// TwinCAT 3 PLC project BottleFactory
// ProgramVersion: 3.1.4026.28
// libraries:
//   CNM_AbstractObject, * (ekvip automation GmbH)
//   CNM_AssertionInterfaces, * (ekvip automation GmbH)
//   CNM_CommandInterfaces, * (ekvip automation GmbH)
//   CNM_CycleManager, * (ekvip automation GmbH)
//   CNM_CycleManagerInterfaces, * (ekvip automation GmbH)
//   CNM_MessageInterfaces, * (ekvip automation GmbH)
//   CNM_ReturnTypes, * (ekvip automation GmbH)
//   CNM_UnicodeUtilities, * (ekvip automation GmbH)
//   Tc2_Standard, * (Beckhoff Automation GmbH)
//   Tc2_System, * (Beckhoff Automation GmbH)
// project tree:
//   / PlcTask.TcTTO
//   POUs/ FB_CappingStation.TcPOU, FB_CinnamonFillingStation.TcPOU, FB_FillingStation.TcPOU, MAIN.TcPOU
// real-time tasks:
//   TASK PlcTask: cycle T#10ms, priority 20, ADS port 350

CONFIGURATION BottleFactory
    RESOURCE PLC ON TwinCAT3
        TASK PlcTask(INTERVAL := T#10ms, PRIORITY := 20);
        PROGRAM MAIN WITH PlcTask : MAIN;
    END_RESOURCE
END_CONFIGURATION

// ---- POUs/MAIN.TcPOU

PROGRAM MAIN
VAR
    bStart : BOOL := FALSE;
    bStop : BOOL := FALSE;
    bBottlePresent : BOOL := TRUE;

    fbStation : FB_FillingStation;
	fbCinnamon : FB_CinnamonFillingStation;
	bCinnamonRun : BOOL := FALSE;
	bCinnamonStop : BOOL := FALSE;
    nConveyorPosition : UDINT;
    nConveyorIndexBase : UDINT;
    nTransferPhase : UDINT;
    nPlaceProgress : UDINT;
    bBottleCapped : BOOL;
    fbInfeed : TON;
    fbOutfeed : TON;
    fbPlacement : TON;
    fbCapping : FB_CappingStation;
END_VAR


// 0: fill, 1: travel to capper, 2: cap, 3: pick and place, 4: bring next bottle to filler.
fbInfeed(IN := nTransferPhase = 1 AND NOT bCinnamonStop, PT := T#2S);
fbCapping(bBottleReady := nTransferPhase = 2, bStop := bCinnamonStop);
fbPlacement(IN := nTransferPhase = 3 AND NOT bCinnamonStop, PT := T#3S);
fbOutfeed(IN := nTransferPhase = 4 AND NOT bCinnamonStop, PT := T#2S);

IF NOT bCinnamonStop THEN
    CASE nTransferPhase OF
        0: IF fbCinnamon.bDone THEN nTransferPhase := 1; END_IF;
        1: IF fbInfeed.Q THEN nTransferPhase := 2; END_IF;
        2: IF fbCapping.bDone THEN nTransferPhase := 3; END_IF;
        3: IF fbPlacement.Q THEN nTransferPhase := 4; END_IF;
        4:
            IF fbOutfeed.Q THEN
                nConveyorIndexBase := nConveyorIndexBase + UDINT#100;
                nTransferPhase := 0;
            END_IF;
    END_CASE;

    nPlaceProgress := 0;
    nConveyorPosition := nConveyorIndexBase;
    CASE nTransferPhase OF
        1: nConveyorPosition := nConveyorIndexBase + DINT_TO_UDINT(TIME_TO_DINT(fbInfeed.ET) / DINT#40);
        2: nConveyorPosition := nConveyorIndexBase + UDINT#50;
        3:
            nConveyorPosition := nConveyorIndexBase + UDINT#50;
            nPlaceProgress := DINT_TO_UDINT(TIME_TO_DINT(fbPlacement.ET) / DINT#30);
        4:
            nConveyorPosition := nConveyorIndexBase + UDINT#50
                + DINT_TO_UDINT(TIME_TO_DINT(fbOutfeed.ET) / DINT#40);
            nPlaceProgress := 100;
    END_CASE;
END_IF;

bBottlePresent := nTransferPhase = 0;
bBottleCapped := nTransferPhase = 3;

fbStation(
    bStart := bStart,
    bStop := bStop,
    bBottlePresent := bBottlePresent
);


fbCinnamon(
    bRunRequest := bCinnamonRun,
    bStop := bCinnamonStop,
    bBottlePresent := bBottlePresent
);

END_PROGRAM

// ---- POUs/FB_FillingStation.TcPOU

FUNCTION_BLOCK FB_FillingStation
VAR_INPUT
    bStart : BOOL;
    bStop : BOOL;
    bBottlePresent : BOOL;
END_VAR

VAR_OUTPUT
    bValveOpen : BOOL;
    bBusy : BOOL;
    bDone : BOOL;
    nCompleted : UDINT;
END_VAR

VAR
    fbTimer : TON;
    fbStartEdge : R_TRIG;
    nState : INT := 0;
END_VAR


fbStartEdge(CLK := bStart);

fbTimer(
    IN := (nState = 10)
          AND NOT bStop
          AND bBottlePresent,
    PT := T#3S
);

bValveOpen := FALSE;
bBusy := FALSE;
bDone := FALSE;

CASE nState OF

    0: // IDLE
        IF fbStartEdge.Q
           AND bBottlePresent
           AND NOT bStop THEN
            nState := 10;
        END_IF;

    10: // FILLING
        IF bStop OR NOT bBottlePresent THEN
            nState := 0;

        ELSIF fbTimer.Q THEN
            nCompleted := nCompleted + 1;
            bDone := TRUE;
            nState := 20;

        ELSE
            bValveOpen := TRUE;
            bBusy := TRUE;
        END_IF;

    20: // COMPLETE
        bDone := TRUE;

        IF NOT bStart THEN
            nState := 0;
        END_IF;

ELSE
    nState := 0;

END_CASE;

END_FUNCTION_BLOCK

// ---- POUs/FB_CinnamonFillingStation.TcPOU

FUNCTION_BLOCK FB_CinnamonFillingStation
VAR_INPUT
    bRunRequest : BOOL;
    bStop : BOOL;
    bBottlePresent : BOOL;
END_VAR

VAR_OUTPUT
    bValveOpen : BOOL;
    bBusy : BOOL;
    bDone : BOOL;
    nCompleted : UDINT;
    nFillPercent : UDINT;
END_VAR

VAR
    fbCycle : CNM_CycleManager.SimpleCycleManager;
    fbTimer : TON;
    bCounted : BOOL := FALSE;
END_VAR

VAR CONSTANT
    STEP_FILL : DINT := 2;
    FILL_DURATION : TIME := T#8S;
END_VAR


(* Update the cycle manager once per PLC scan *)
fbCycle(
    execute := bRunRequest
               AND bBottlePresent
               AND NOT bStop
);

(* Filling timer *)
fbTimer(
    IN := fbCycle.step.current = STEP_FILL,
    PT := FILL_DURATION
);

(* Default outputs *)
bValveOpen := FALSE;
bBusy := FALSE;
bDone := FALSE;
nFillPercent := 0;

CASE fbCycle.step.current OF

    CNM_ReturnTypes.DefaultSteps.STEP.INIT:
        bCounted := FALSE;
        fbCycle.proceed();

    STEP_FILL:
        bBusy := TRUE;
        nFillPercent := DINT_TO_UDINT(TIME_TO_DINT(fbTimer.ET) * DINT#100 / TIME_TO_DINT(FILL_DURATION));
        bValveOpen := NOT fbTimer.Q;

        fbCycle.step.next :=
            CNM_ReturnTypes.DefaultSteps.STEP.SUCCESS;

        fbCycle.waitFor(value := fbTimer.Q);

    CNM_ReturnTypes.DefaultSteps.STEP.SUCCESS:
        bDone := TRUE;
        nFillPercent := 100;

        IF NOT bCounted THEN
            nCompleted := nCompleted + 1;
            bCounted := TRUE;
        END_IF;

END_CASE;

END_FUNCTION_BLOCK

// ---- POUs/FB_CappingStation.TcPOU

FUNCTION_BLOCK FB_CappingStation
VAR_INPUT
    bBottleReady : BOOL;
    bStop : BOOL;
END_VAR
VAR_OUTPUT
    bDone : BOOL;
    nArmProgress : UDINT;
END_VAR
VAR
    fbCycle : CNM_CycleManager.SimpleCycleManager;
    fbArmTimer : TON;
END_VAR
VAR CONSTANT
    STEP_CAP : DINT := 2;
    ARM_DURATION : TIME := T#2S;
END_VAR


fbCycle(execute := bBottleReady AND NOT bStop);
fbArmTimer(IN := fbCycle.step.current = STEP_CAP AND bBottleReady AND NOT bStop,
           PT := ARM_DURATION);

bDone := FALSE;
nArmProgress := 0;

IF bBottleReady AND NOT bStop THEN
    CASE fbCycle.step.current OF
        CNM_ReturnTypes.DefaultSteps.STEP.INIT:
            fbCycle.proceed();

        STEP_CAP:
            nArmProgress := DINT_TO_UDINT(TIME_TO_DINT(fbArmTimer.ET) * DINT#100
                                          / TIME_TO_DINT(ARM_DURATION));
            fbCycle.step.next := CNM_ReturnTypes.DefaultSteps.STEP.SUCCESS;
            fbCycle.waitFor(value := fbArmTimer.Q);

        CNM_ReturnTypes.DefaultSteps.STEP.SUCCESS:
            nArmProgress := 100;
            bDone := TRUE;
    END_CASE;
END_IF;

END_FUNCTION_BLOCK
